ABB RAPID module: LabJointRws.mod

MODULE LabJointRws
  ! V5 servidor PC (20/11/2026). Docs: rws_mover.py. Max 5000 caracteres.
  ! PC escribe pcTarget (+pcTipo/pcPose), lo relee y sube pcSeq. Robot valida,
  ! mueve con fine, publica rbCodigo y luego rbSeq. pcTipo 0 MoveAbsJ pcTarget,
  ! 1 MoveL pcPose (tool0, wobj0). rbCodigo 1 moviendo 2 llegada -1 vacio
  ! -2 limites -3 paso -4 modo -5 tipo.
  CONST num maxPasoDeg := 360;
  CONST num margenDeg := 2;
  CONST bool permitirAuto := FALSE;
  CONST speeddata vMax := [250,60,250,60];
  PERS num pcVelPct := 20;
  PERS jointtarget pcTarget := [[9E9,9E9,9E9,9E9,9E9,9E9],[9E9,9E9,9E9,9E9,9E9,9E9]];
  PERS num pcTipo := 0;
  PERS robtarget pcPose := [[9E9,9E9,9E9],[1,0,0,0],[0,0,0,0],[9E9,9E9,9E9,9E9,9E9,9E9]];
  PERS num pcSeq := 0;
  PERS num pcFin := 0;
  PERS num rbSeq := 0;
  PERS num rbCodigo := 0;
  PERS num rbActivo := 0;

  PROC MostrarObjetivo()
    MostrarEjes pcTarget.robax;
  ENDPROC

  PROC ServidorPC()
    VAR jointtarget objetivo;
    VAR jointtarget actual;
    VAR robtarget destino;
    VAR num tipo := 0;
    VAR num seq := 0;
    VAR num respuesta := 0;
    VAR errnum motivo := 0;
    VAR speeddata vOrden;
    VAR num pct := 20;

    rbActivo := 0;
    IF ModoPermitido() = FALSE THEN
      TPWrite "Seleccione manual reducido.";
      RETURN;
    ENDIF
    TPReadFK respuesta,"Aceptar objetivos enviados por la PC?",stEmpty,stEmpty,stEmpty,"Iniciar","Cancelar"\MaxTime:=120\BreakFlag:=motivo;
    IF motivo <> 0 OR respuesta <> 4 THEN
      TPWrite "Servidor PC cancelado.";
      RETURN;
    ENDIF
    pcFin := 0;
    rbCodigo := 0;
    rbSeq := pcSeq;
    rbActivo := 1;
    AccSet 50, 50;
    TPWrite "Servidor PC activo. Esperando objetivos.";
    WHILE pcFin = 0 DO
      IF pcSeq <> rbSeq THEN
        seq := pcSeq;
        objetivo := pcTarget;
        tipo := pcTipo;
        destino := pcPose;
        actual := CJointT();
        rbCodigo := Validar(objetivo.robax, actual.robax, tipo, destino);
        IF rbCodigo = 0 THEN
          rbCodigo := 1;
          TPWrite "Moviendo orden"\Num:=seq;
          objetivo.extax := actual.extax;
          pct := pcVelPct;
          IF pct < 1 OR pct > 100 THEN
            pct := 20;
          ENDIF
          vOrden := vMax;
          vOrden.v_tcp := vMax.v_tcp * pct / 100;
          vOrden.v_ori := vMax.v_ori * pct / 100;
          IF tipo = 0 THEN
            MoveAbsJ objetivo,vOrden,fine,tool0;
          ELSE
            ConfL\Off;
            MoveL destino,vOrden,fine,tool0\WObj:=wobj0;
            ConfL\On;
          ENDIF
          rbCodigo := 2;
        ELSE
          TPWrite "Orden rechazada, codigo"\Num:=rbCodigo;
        ENDIF
        rbSeq := seq;
      ENDIF
      WaitTime 0.1;
    ENDWHILE
    rbActivo := 0;
    AccSet 100, 100;
    TPWrite "Servidor PC terminado.";
  ENDPROC

  LOCAL PROC MostrarEjes(robjoint ejes)
    TPWrite "Objetivo absoluto en grados:";
    TPWrite "J1"\Num:=ejes.rax_1;
    TPWrite "J2"\Num:=ejes.rax_2;
    TPWrite "J3"\Num:=ejes.rax_3;
    TPWrite "J4"\Num:=ejes.rax_4;
    TPWrite "J5"\Num:=ejes.rax_5;
    TPWrite "J6"\Num:=ejes.rax_6;
  ENDPROC

  LOCAL FUNC bool ModoPermitido()
    VAR bool permitido := FALSE;
    IF OpMode() = OP_MAN_PROG THEN
      permitido := TRUE;
    ELSEIF permitirAuto THEN
      IF OpMode() = OP_AUTO THEN
        permitido := TRUE;
      ENDIF
    ENDIF
    RETURN permitido;
  ENDFUNC

  LOCAL FUNC num Validar(robjoint q, robjoint actual, num tipo, robtarget p)
    IF ModoPermitido() = FALSE THEN
      RETURN -4;
    ENDIF
    IF tipo <> 0 AND tipo <> 1 THEN
      RETURN -5;
    ENDIF
    IF tipo = 1 AND (Abs(p.trans.x) > 2000 OR Abs(p.trans.y) > 2000 OR
     Abs(p.trans.z) > 2000) THEN
      RETURN -1;
    ENDIF
    IF Abs(q.rax_1) > 1000 OR Abs(q.rax_2) > 1000 OR Abs(q.rax_3) > 1000 OR
     Abs(q.rax_4) > 1000 OR Abs(q.rax_5) > 1000 OR Abs(q.rax_6) > 1000 THEN
      RETURN -1;
    ENDIF
    IF q.rax_1 < (-165 + margenDeg) OR q.rax_1 > (165 - margenDeg) OR
     q.rax_2 < (-110 + margenDeg) OR q.rax_2 > (110 - margenDeg) OR
     q.rax_3 < (-110 + margenDeg) OR q.rax_3 > (70 - margenDeg) OR
     q.rax_4 < (-160 + margenDeg) OR q.rax_4 > (160 - margenDeg) OR
     q.rax_5 < (-120 + margenDeg) OR q.rax_5 > (120 - margenDeg) OR
     q.rax_6 < (-400 + margenDeg) OR q.rax_6 > (400 - margenDeg) THEN
      RETURN -2;
    ENDIF
    IF Abs(q.rax_1 - actual.rax_1) > maxPasoDeg OR Abs(q.rax_2 - actual.rax_2) > maxPasoDeg OR
     Abs(q.rax_3 - actual.rax_3) > maxPasoDeg OR Abs(q.rax_4 - actual.rax_4) > maxPasoDeg OR
     Abs(q.rax_5 - actual.rax_5) > maxPasoDeg OR Abs(q.rax_6 - actual.rax_6) > maxPasoDeg THEN
      RETURN -3;
    ENDIF
    RETURN 0;
  ENDFUNC
ENDMODULE
